(* IEC 61131-3 sources: trust-platform/examples/OSCAT/mixed_vendor_vfd_adapter/non-oop/src, 3 files *)

(* ---- Main.st ---- *)
FUNCTION_BLOCK ClassicMotorCell
VAR
    RunningCountValue : INT;
    FaultCountValue : INT;
    LastFaultCodeValue : DWORD;
END_VAR

METHOD PUBLIC Update : INT
VAR_INPUT
    AbbStatus : WORD;
    DanfossStatus : WORD;
    SiemensStatus : WORD;
    RunCommand : BOOL;
    PullCordOk : BOOL;
END_VAR
RunningCountValue := INT#0;
FaultCountValue := INT#0;
LastFaultCodeValue := DWORD#0;
IF PullCordOk AND RunCommand THEN
    IF (WORD_TO_DWORD(AbbStatus) AND DWORD#16#0004) <> DWORD#0 THEN
        RunningCountValue := RunningCountValue + INT#1;
    END_IF;
    IF (WORD_TO_DWORD(AbbStatus) AND DWORD#16#0008) <> DWORD#0 THEN
        FaultCountValue := FaultCountValue + INT#1;
        LastFaultCodeValue := DWORD#16#10000011;
    END_IF;
    IF (WORD_TO_DWORD(DanfossStatus) AND DWORD#16#0100) <> DWORD#0 THEN
        RunningCountValue := RunningCountValue + INT#1;
    END_IF;
    IF (WORD_TO_DWORD(DanfossStatus) AND DWORD#16#0002) <> DWORD#0 THEN
        FaultCountValue := FaultCountValue + INT#1;
        LastFaultCodeValue := DWORD#16#20000022;
    END_IF;
    IF (WORD_TO_DWORD(SiemensStatus) AND DWORD#16#0400) <> DWORD#0 THEN
        RunningCountValue := RunningCountValue + INT#1;
    END_IF;
    IF (WORD_TO_DWORD(SiemensStatus) AND DWORD#16#0008) <> DWORD#0 THEN
        FaultCountValue := FaultCountValue + INT#1;
        LastFaultCodeValue := DWORD#16#30000033;
    END_IF;
END_IF;
Update := FaultCountValue;
END_METHOD

PUBLIC PROPERTY RunningCount : INT
GET
    RunningCount := RunningCountValue;
END_GET
END_PROPERTY

PUBLIC PROPERTY LastFaultCode : DWORD
GET
    LastFaultCode := LastFaultCodeValue;
END_GET
END_PROPERTY
END_FUNCTION_BLOCK

PROGRAM Main
VAR
    Cell : ClassicMotorCell;
    Faults : INT;
END_VAR
Faults := Cell.Update(AbbStatus := WORD#16#0004, DanfossStatus := WORD#16#0100, SiemensStatus := WORD#16#0400, RunCommand := TRUE, PullCordOk := TRUE);
END_PROGRAM

(* ---- Configuration.st ---- *)
CONFIGURATION MixedVendorVfdAdapterClassicConfiguration
RESOURCE Cpu0 ON PLC
    TASK MainTask (INTERVAL := T#100ms, PRIORITY := 1);
    PROGRAM Cell WITH MainTask : Main;
END_RESOURCE
END_CONFIGURATION

(* ---- Tests.st ---- *)
TEST_PROGRAM ClassicMotorCellDecodesVendorBitsInline
VAR
    Cell : ClassicMotorCell;
END_VAR

ASSERT_EQUAL(EXPECTED := INT#1, ACTUAL := Cell.Update(AbbStatus := WORD#16#0004, DanfossStatus := WORD#16#0002, SiemensStatus := WORD#16#0400, RunCommand := TRUE, PullCordOk := TRUE));
ASSERT_EQUAL(EXPECTED := DWORD#16#20000022, ACTUAL := Cell.LastFaultCode);
END_TEST_PROGRAM
